Staubli VAL3: moveCalPos.pgx

program moveCalPos(string x_sTarget)
  local bool l_bTaskStatusErr
begin
  if taskStatus("m")!=-1
    taskKill("m")
  endIf
  if taskStatus("m")==-1
    taskCreate "m",100, db:ListMove(x_sTarget)
  endIf
  l_bTaskStatusErr=watch(taskStatus("m")==150 or taskStatus("m")>1,0.3)
  if l_bTaskStatusErr==true
    taskKill("m")
    call db:hmiAlert("CantMove1","warning")
  endIf
end
